Fanuc KAREL source: kc00061.KL

-- PROVISIONAL review KL for V1013-1; original PC SHA256 ac0e36d82a02f80339886f28752c7048bdbea91d0b6910914b3ca6e8275148ef
-- Incomplete behavior may be omitted. Consult companion uncertainty JSON. Do not deploy.
PROGRAM KC00061
%NOLOCKGROUP
BEGIN
  -- UNRESOLVED_PC offsets 5-37; opcodes 27,27,9D,27,9D,22,1C,22,AA,23
  -- UNRESOLVED_PC offsets 42-46; opcodes 7F
END KC00061
